ORGANIZATION_BLOCK "Main"
{ S7_Optimized_Access := 'TRUE' }
VERSION : 0.1
BEGIN
   "Result" := "Calculate"(X := 5.0);
END_ORGANIZATION_BLOCK
